Fanuc KAREL source: KC00039.KL

PROGRAM KC00039
%NOLOCKGROUP
VAR
  I: INTEGER
  J: INTEGER
  K: INTEGER
  R: REAL
  B: BOOLEAN
  S: STRING[80]
  T: STRING[80]
  P: PATH
  Q: PATH
  AI: ARRAY[8] OF INTEGER
  AB: ARRAY[244] OF BYTE
  JP: JOINTPOS
  AR: ARRAY[9] OF REAL
BEGIN
  CNV_REL_JPOS(AR,JP,I)
END KC00039
